Fanuc KAREL source: KO00062.KL

PROGRAM KO00062
%NOLOCKGROUP
%ENVIRONMENT MIR
VAR
  P1: XYZWPR
  P2: JOINTPOS
  F: BOOLEAN
  OUT: XYZWPR
BEGIN
  F = TRUE
  OUT = MIRROR(P1, P2, F)
END KO00062
